{region 'Documentation'}
(*!
<summary>Delays only the concrete Reset completion; all lifecycle and reservation processing remains inherited.</summary>
*)
{endregion}
FUNCTION_BLOCK ReservationResetChild EXTENDS ReservationChildProbe
VAR_INPUT
    AllowResetCompletion : BOOL := TRUE; //! FALSE holds the real child in Reset; TRUE permits inherited Reset completion.
END_VAR

SUPER^();

{region 'Documentation'}
(*!
<summary>Completes the concrete Reset only when released by the local scenario.</summary>
*)
{endregion}
METHOD PROTECTED ProcessReset
IF AllowResetCompletion THEN
    SUPER^.ProcessReset();
END_IF;
END_METHOD

END_FUNCTION_BLOCK

(* stored: Version 1.1.0.1
   POU ReservationResetChild: Id {b4ae866e-452a-4984-bc65-f40f6ac0cc58}, SpecialFunc None
   Folder Internal: Id {b4bebbf7-61eb-417e-a45b-083a3c14a85c}
   Method ProcessReset: Id {fa04e567-55e6-4011-a95f-530ccfbc72ae} *)
